Fanuc KAREL source: KT00350.KL

PROGRAM KT00350
%NOLOCKGROUP
VAR
  P1: POSITION
  P2: JOINTPOS
  OUT: BOOLEAN
BEGIN
  OUT = P1 < P2
END KT00350
